(* IEC 61131-3 sources: axsharp/src/tests.integrations/integrated/src/ax/src, 2 files *)

(* ---- configuration.st ---- *)
USING RealMonsterData;
CONFIGURATION MyConfiguration
    TASK Main(Interval := T#10ms, Priority := 1);
    PROGRAM P1 WITH Main: MyProgram;

    VAR_GLOBAL
       {S7.extern=ReadWrite}
       Monster : MonsterData.Monster;
       {S7.extern=ReadWrite}
       OnlineToPlain_should_copy_entire_structure : MonsterData.Monster;
       {S7.extern=ReadWrite}
       PlainToOnline_should_copy_entire_structure : MonsterData.Monster;
       {S7.extern=ReadWrite}
       OnlineToShadowAsync_should_copy_entire_structure : MonsterData.Monster;
       {S7.extern=ReadWrite}
       ShadowToOnlineAsync_should_copy_entire_structure : MonsterData.Monster;

       {S7.extern=ReadWrite}
       ITwinObjectOnlineToPlain_should_copy_entire_structure : MonsterData.Monster;
       {S7.extern=ReadWrite}
       ITwinObjectPlainToOnline_should_copy_entire_structure : MonsterData.Monster;
       {S7.extern=ReadWrite}
       ITwinObjectOnlineToShadowAsync_should_copy_entire_structure : MonsterData.Monster;
       {S7.extern=ReadWrite}
       ITwinObjectShadowToOnlineAsync_should_copy_entire_structure : MonsterData.Monster;

       {S7.extern=ReadWrite}
       ShadowToPlainAsync_should_copy_entire_structure : MonsterData.Monster;
       {S7.extern=ReadWrite}
       PlainToShadowAsync_should_copy_entire_structure : MonsterData.Monster;

       {S7.extern=ReadWrite}
       ITwinObjectShadowToPlainAsync_should_copy_entire_structure : MonsterData.Monster;
       {S7.extern=ReadWrite}
       ITwinObjectPlainToShadowAsync_should_copy_entire_structure : MonsterData.Monster;

       {S7.extern=ReadWrite}
       Pokus : Pokus;

       {S7.extern=ReadWrite}
       RealMonster : RealMonsterData.RealMonster;
       {S7.extern=ReadWrite}
       OnlineToShadow_should_copy : RealMonsterData.RealMonster;
       {S7.extern=ReadWrite}
       ShadowToOnline_should_copy : RealMonsterData.RealMonster;
       {S7.extern=ReadWrite}
       OnlineToPlain_should_copy: RealMonsterData.RealMonster;
       {S7.extern=ReadWrite}
       PlainToOnline_should_copy: RealMonsterData.RealMonster;

       {S7.extern=ReadWrite}
       ITwinObjectOnlineToShadow_should_copy : RealMonsterData.RealMonster;
       {S7.extern=ReadWrite}
       ITwinObjectShadowToOnline_should_copy : RealMonsterData.RealMonster;
       {S7.extern=ReadWrite}
       ITwinObjectOnlineToPlain_should_copy: RealMonsterData.RealMonster;
       {S7.extern=ReadWrite}
       ITwinObjectPlainToOnline_should_copy: RealMonsterData.RealMonster;

       {S7.extern=ReadWrite}
       p_online_shadow: all_primitives;
       {S7.extern=ReadWrite}
       p_shadow_online: all_primitives;

       {S7.extern=ReadWrite}
       p_online_plain: all_primitives;
       {S7.extern=ReadWrite}
       p_plain_online: all_primitives;

       {S7.extern=ReadWrite}
       p_shadow_plain: all_primitives;
       {S7.extern=ReadWrite}
       p_plain_shadow: all_primitives;

       {S7.extern=ReadWrite}
       StartPolling_should_update_cyclic_property : RealMonsterData.RealMonster;

       {S7.extern=ReadWrite}
       StartPolling_ConcurentOverload : RealMonsterData.RealMonster;

       {S7.extern=ReadWrite}
       ChangeDetections : RealMonsterData.RealMonster;

       {S7.extern=ReadWrite}
       GH_ISSUE_183 : GH_ISSUE_183.GH_ISSUE_183_1;
    END_VAR
END_CONFIGURATION

CLASS Pokus
    VAR PUBLIC
        Nested : Nested;
    END_VAR

END_CLASS

CLASS Nested
    VAR PUBLIC
        SomeString : STRING;
        SomeInt : INT;
        SomeByte : BYTE;
    END_VAR
END_CLASS

(* ---- program.st ---- *)
PROGRAM MyProgram
    VAR_EXTERNAL
        StartPolling_should_update_cyclic_property : RealMonsterData.RealMonster;
        GH_ISSUE_183 : GH_ISSUE_183.GH_ISSUE_183_1;

        StartPolling_ConcurentOverload : RealMonsterData.RealMonster;
    END_VAR
    StartPolling_should_update_cyclic_property.Id := StartPolling_should_update_cyclic_property.Id + ULINT#1;

    StartPolling_should_update_cyclic_property.DriveA.NestedLevelOne.NestedLevelTwo.NestedLevelThree.Position := StartPolling_should_update_cyclic_property.DriveA.NestedLevelOne.NestedLevelTwo.NestedLevelThree.Position  + REAL#1.0;

    StartPolling_ConcurentOverload.Id := StartPolling_ConcurentOverload.Id + ULINT#1;

    StartPolling_ConcurentOverload.ArrayOfBytes[0] := StartPolling_ConcurentOverload.ArrayOfBytes[1];
    StartPolling_ConcurentOverload.ArrayOfBytes[1] := StartPolling_ConcurentOverload.ArrayOfBytes[2];
    StartPolling_ConcurentOverload.ArrayOfBytes[2] := StartPolling_ConcurentOverload.ArrayOfBytes[3];
    StartPolling_ConcurentOverload.ArrayOfBytes[3] := TO_BYTE( TO_INT(StartPolling_ConcurentOverload.ArrayOfBytes[0]) + 1 );

    StartPolling_ConcurentOverload.ArrayOfDrives[0].Position    := StartPolling_ConcurentOverload.ArrayOfDrives[1].Position ;
    StartPolling_ConcurentOverload.ArrayOfDrives[0].Velo        := StartPolling_ConcurentOverload.ArrayOfDrives[1].Velo ;
    StartPolling_ConcurentOverload.ArrayOfDrives[0].Dcc         := StartPolling_ConcurentOverload.ArrayOfDrives[1].Acc ;
    StartPolling_ConcurentOverload.ArrayOfDrives[0].Acc         := StartPolling_ConcurentOverload.ArrayOfDrives[1].Dcc ;

    StartPolling_ConcurentOverload.ArrayOfDrives[1].Position    := StartPolling_ConcurentOverload.ArrayOfDrives[2].Position ;
    StartPolling_ConcurentOverload.ArrayOfDrives[1].Velo        := StartPolling_ConcurentOverload.ArrayOfDrives[2].Velo ;
    StartPolling_ConcurentOverload.ArrayOfDrives[1].Dcc         := StartPolling_ConcurentOverload.ArrayOfDrives[2].Acc ;
    StartPolling_ConcurentOverload.ArrayOfDrives[1].Acc         := StartPolling_ConcurentOverload.ArrayOfDrives[2].Dcc ;

    StartPolling_ConcurentOverload.ArrayOfDrives[2].Position    := StartPolling_ConcurentOverload.ArrayOfDrives[3].Position ;
    StartPolling_ConcurentOverload.ArrayOfDrives[2].Velo        := StartPolling_ConcurentOverload.ArrayOfDrives[3].Velo ;
    StartPolling_ConcurentOverload.ArrayOfDrives[2].Dcc         := StartPolling_ConcurentOverload.ArrayOfDrives[3].Acc ;
    StartPolling_ConcurentOverload.ArrayOfDrives[2].Acc         := StartPolling_ConcurentOverload.ArrayOfDrives[3].Dcc ;

    StartPolling_ConcurentOverload.ArrayOfDrives[3].Position    := StartPolling_ConcurentOverload.ArrayOfDrives[0].Position + 0.02;
    StartPolling_ConcurentOverload.ArrayOfDrives[3].Velo        := StartPolling_ConcurentOverload.ArrayOfDrives[0].Velo + 0.03;
    StartPolling_ConcurentOverload.ArrayOfDrives[3].Dcc         := StartPolling_ConcurentOverload.ArrayOfDrives[0].Acc + 0.04;
    StartPolling_ConcurentOverload.ArrayOfDrives[3].Acc         := StartPolling_ConcurentOverload.ArrayOfDrives[0].Dcc + 0.05;

    StartPolling_ConcurentOverload.DriveA.Position    := StartPolling_ConcurentOverload.ArrayOfDrives[0].Position ;
    StartPolling_ConcurentOverload.DriveA.Velo        := StartPolling_ConcurentOverload.ArrayOfDrives[0].Velo ;
    StartPolling_ConcurentOverload.DriveA.Dcc         := StartPolling_ConcurentOverload.ArrayOfDrives[0].Acc ;
    StartPolling_ConcurentOverload.DriveA.Acc         := StartPolling_ConcurentOverload.ArrayOfDrives[0].Dcc ;

    StartPolling_ConcurentOverload.DriveA.NestedLevelOne.Position    := StartPolling_ConcurentOverload.ArrayOfDrives[1].Position ;
    StartPolling_ConcurentOverload.DriveA.NestedLevelOne.Velo        := StartPolling_ConcurentOverload.ArrayOfDrives[1].Velo ;
    StartPolling_ConcurentOverload.DriveA.NestedLevelOne.Dcc         := StartPolling_ConcurentOverload.ArrayOfDrives[1].Acc ;
    StartPolling_ConcurentOverload.DriveA.NestedLevelOne.Acc         := StartPolling_ConcurentOverload.ArrayOfDrives[1].Dcc ;

    StartPolling_ConcurentOverload.DriveA.NestedLevelOne.NestedLevelTwo.Position    := StartPolling_ConcurentOverload.ArrayOfDrives[2].Position ;
    StartPolling_ConcurentOverload.DriveA.NestedLevelOne.NestedLevelTwo.Velo        := StartPolling_ConcurentOverload.ArrayOfDrives[2].Velo ;
    StartPolling_ConcurentOverload.DriveA.NestedLevelOne.NestedLevelTwo.Dcc         := StartPolling_ConcurentOverload.ArrayOfDrives[2].Acc ;
    StartPolling_ConcurentOverload.DriveA.NestedLevelOne.NestedLevelTwo.Acc         := StartPolling_ConcurentOverload.ArrayOfDrives[2].Dcc ;

    StartPolling_ConcurentOverload.DriveA.NestedLevelOne.NestedLevelTwo.NestedLevelThree.Position    := StartPolling_ConcurentOverload.ArrayOfDrives[3].Position ;
    StartPolling_ConcurentOverload.DriveA.NestedLevelOne.NestedLevelTwo.NestedLevelThree.Velo        := StartPolling_ConcurentOverload.ArrayOfDrives[3].Velo ;
    StartPolling_ConcurentOverload.DriveA.NestedLevelOne.NestedLevelTwo.NestedLevelThree.Dcc         := StartPolling_ConcurentOverload.ArrayOfDrives[3].Acc ;
    StartPolling_ConcurentOverload.DriveA.NestedLevelOne.NestedLevelTwo.NestedLevelThree.Acc         := StartPolling_ConcurentOverload.ArrayOfDrives[3].Dcc ;

END_PROGRAM
